FUNCTION_BLOCK FallbackElapsedTimeCtrl (* Basic Function Block Type *)
  (* Standard: 61499-2 *)
  (* Version 0.0, 10/7/2026, Schneider Electric, Template *)
  PACKAGE SE.Nereda;
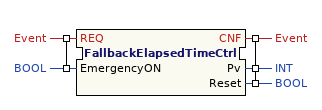
  EVENT_INPUT
    REQ WITH EmergencyON; (* Normal Execution Request *)
  END_EVENT
  EVENT_OUTPUT
    CNF WITH Pv, Reset; (* Execution Confirmation *)
  END_EVENT
  VAR_INPUT
    EmergencyON : BOOL; (* Input event qualifier *)
  END_VAR
  VAR_OUTPUT
    Pv : INT; (* Output event qualifier *)
    Reset : BOOL;
  END_VAR
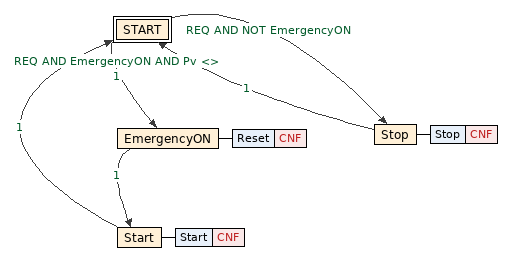
  EC_STATES
    START; (* Initial State *)
    EmergencyON : Reset -> CNF;
    Start : Start -> CNF;
    Stop : Stop -> CNF;
  END_STATES
  EC_TRANSITIONS
    START TO EmergencyON := REQ AND EmergencyON AND Pv <> 1;
    EmergencyON TO Start := 1;
    Start TO START := 1;
    START TO Stop := REQ AND NOT EmergencyON;
    Stop TO START := 1;
  END_TRANSITIONS
  ALGORITHM Reset IN ST:
;
Reset := TRUE;
  END_ALGORITHM
  ALGORITHM Start IN ST:
;
Pv := 1;
Reset := FALSE;
  END_ALGORITHM
  ALGORITHM Stop IN ST:
;
Pv := 0;
Reset := FALSE;
  END_ALGORITHM
END_FUNCTION_BLOCK
